(* IEC 61131-3 sources: rusty/tests/lit/cfc/blocks/function_call, 2 files *)

(* ---- main.st ---- *)
FUNCTION main : DINT
    VAR
        result : DINT;
        doubled : DINT;
    END_VAR
    result := function_call(in1 := 3, in2 := 4, doubledOut => doubled);
    // CHECK: result = 7, doubled = 14
    printf('result = %d, doubled = %d$N', result, doubled);
END_FUNCTION

(* ---- myAdd.st ---- *)
FUNCTION myAdd : INT
    VAR_INPUT
        in1, in2: DINT;
    END_VAR

    VAR_OUTPUT
        myAddDoubled: DINT;
    END_VAR

    myAdd := in1 + in2;
    myAddDoubled := (in1 + in2) * 2;
END_FUNCTION
